(* LS Electric XG5000 project: Crane11 *)
(* PLC LSPLC *)
(* module base 0 slot 0: 입출력 모듈:XGH-DT4A (DC 24V 입력, 트랜지스터 출력 32점 ) *)
(* module base 0 slot 1: Cnet:XGL-C42A/B (Cnet 통신 모듈(RS-422/485, RS-422/485)) *)
VAR_GLOBAL
    AUTO_MODE_1 AT %IX0.0.0 : BOOL;
    AUTO_MODE_2 AT %IX0.0.1 : BOOL;
    AUTO_POSITION AT %IX0.0.6 : BOOL;
    AUTO_RESET AT %IX0.0.4 : BOOL;
    AUTO_RESUME AT %IX0.0.5 : BOOL;
    AUTO_START AT %IX0.0.2 : BOOL;
    AUTO_STOP AT %IX0.0.3 : BOOL;
    DRV_VAL AT %MW1 : WORD;
    DRV_VAL_GLOBAL : WORD;
    FREQ_VAL AT %MW0 : WORD;
    FREQ_VAL_GLOBAL : WORD;
    HALL_SENSOR_RPM AT %IX0.0.11 : BOOL;
    LED_AUTO_POSITION AT %QX0.0.19 : BOOL;
    LED_AUTO_RESET AT %QX0.0.20 : BOOL;
    LED_AUTO_RESUME AT %QX0.0.18 : BOOL;
    LED_AUTO_START AT %QX0.0.16 : BOOL;
    LED_AUTO_STOP AT %QX0.0.17 : BOOL;
    LIMITE_SW_BOTTOM_LEFT AT %IX0.0.13 : BOOL;
    LIMITE_SW_BOTTOM_RIGHT AT %IX0.0.15 : BOOL;
    LIMITE_SW_TOP_LEFT AT %IX0.0.12 : BOOL;
    LIMITE_SW_TOP_RIGHT AT %IX0.0.14 : BOOL;
    MODE_SELECT_AUTO AT %IX0.0.9 : BOOL;
    MODE_SELECT_PASSIVE AT %IX0.0.10 : BOOL;
    STATE_AUTO_MODE_1 : BOOL;
    STATE_AUTO_MODE_2 : BOOL;
    STATE_LIMITE_SW_BOTTOM_LEFT : BOOL;
    STATE_LIMITE_SW_BOTTOM_RIGHT : BOOL;
    STATE_POSITION : BOOL;
    STATE_RESET : BOOL;
    STATE_RESUME : BOOL;
    STATE_START : BOOL;
    STATE_STOP : BOOL;
    STATE_STOP_EMERGENCY : BOOL;
    STOP_EMERGENCY AT %IX0.0.7 : BOOL;
    SUCCESS_POSITION : BOOL;
    SUCCESS_RESET : BOOL;
    VAL_STATE_RESET : BOOL;
END_VAR

FUNCTION_BLOCK FB_LED_FLASH
(* 램프 점멸 동작 *)
VAR_INPUT
    EN_SW : BOOL;
    T_ON : TIME;
    T_OFF : TIME;
END_VAR
VAR_OUTPUT
    OUT_LAMP : BOOL;
END_VAR
VAR
    TIMER_1 : TON;
    TIMER_2 : TON;
END_VAR
(* 1. TIMER_1 동작: 시작 스위치가 켜져 있고, TIMER_2가 꺼져있을 때(.Q가 아닐 때) *)
TIMER_1(IN := EN_SW AND NOT TIMER_2.Q, PT := T_ON);

(* 2. TIMER_2 동작: TIMER_1이 완료되었을 때(.Q 일 때) *)
TIMER_2(IN := TIMER_1.Q, PT := T_OFF);

(* 3. 램프 출력: 스위치 ON 상태이고, TIMER_1이 도는 동안(아직 .Q가 안 떴을 때) *)
IF EN_SW AND NOT TIMER_1.Q THEN
    OUT_LAMP := TRUE;
ELSE
    OUT_LAMP := FALSE;
END_IF;
END_FUNCTION_BLOCK

FUNCTION_BLOCK FB_SELF_HOLD
VAR_INPUT
    START_SW : BOOL;
    STOP_SW : BOOL;
END_VAR
VAR_OUTPUT
    MOTOR_START : BOOL;
    MOTOR_STOP : BOOL;
END_VAR
IF STOP_SW THEN
    MOTOR_START := FALSE; // 실제 출력 변수 직접 제어
    MOTOR_STOP  := TRUE;
ELSIF START_SW THEN
    MOTOR_START := TRUE;
    MOTOR_STOP  := FALSE;
END_IF;
END_FUNCTION_BLOCK

PROGRAM LED_OUTPUT (* task: 스캔 프로그램 *)
(* LED출력관련 *)
VAR_EXTERNAL
    AUTO_POSITION : BOOL; (* AT %IX0.0.6 *)
    AUTO_RESET : BOOL; (* AT %IX0.0.4 *)
    AUTO_RESUME : BOOL; (* AT %IX0.0.5 *)
    AUTO_START : BOOL; (* AT %IX0.0.2 *)
    AUTO_STOP : BOOL; (* AT %IX0.0.3 *)
    LED_AUTO_POSITION : BOOL; (* AT %QX0.0.19 *)
    LED_AUTO_RESET : BOOL; (* AT %QX0.0.20 *)
    LED_AUTO_RESUME : BOOL; (* AT %QX0.0.18 *)
    LED_AUTO_START : BOOL; (* AT %QX0.0.16 *)
    LED_AUTO_STOP : BOOL; (* AT %QX0.0.17 *)
    STATE_POSITION : BOOL;
    STATE_RESET : BOOL;
    STATE_RESUME : BOOL;
    STATE_START : BOOL;
    STATE_STOP : BOOL;
    STATE_STOP_EMERGENCY : BOOL;
    STOP_EMERGENCY : BOOL; (* AT %IX0.0.7 *)
    SUCCESS_POSITION : BOOL;
    SUCCESS_RESET : BOOL;
END_VAR
VAR
    AUTO_RESET_STATE : BOOL;
    AUTO_STOP_STATE : BOOL;
    HOLD_EMERGENCY : FB_SELF_HOLD;
    HOLD_POSITION : FB_SELF_HOLD;
    HOLD_POSITION1 : FB_SELF_HOLD;
    HOLD_RESET : FB_SELF_HOLD;
    HOLD_RESET1 : FB_SELF_HOLD;
    HOLD_RESET2 : FB_SELF_HOLD;
    HOLD_START : FB_SELF_HOLD;
    HOLD_START1 : FB_SELF_HOLD;
    HOLD_START2 : FB_SELF_HOLD;
    HOLD_START3 : FB_SELF_HOLD;
    HOLD_STOP : FB_SELF_HOLD;
    LAMP_POSITION : FB_LED_FLASH;
    LAMP_RESET : FB_LED_FLASH;
    LAMP_RESUME : FB_LED_FLASH;
    LOCAL_POSITION : BOOL;
    LOCAL_RESET : BOOL;
    LOCAL_STOP_EMERGENCY : BOOL;
    RESET_STATE : BOOL;
    VAL_STATE : BOOL;
END_VAR

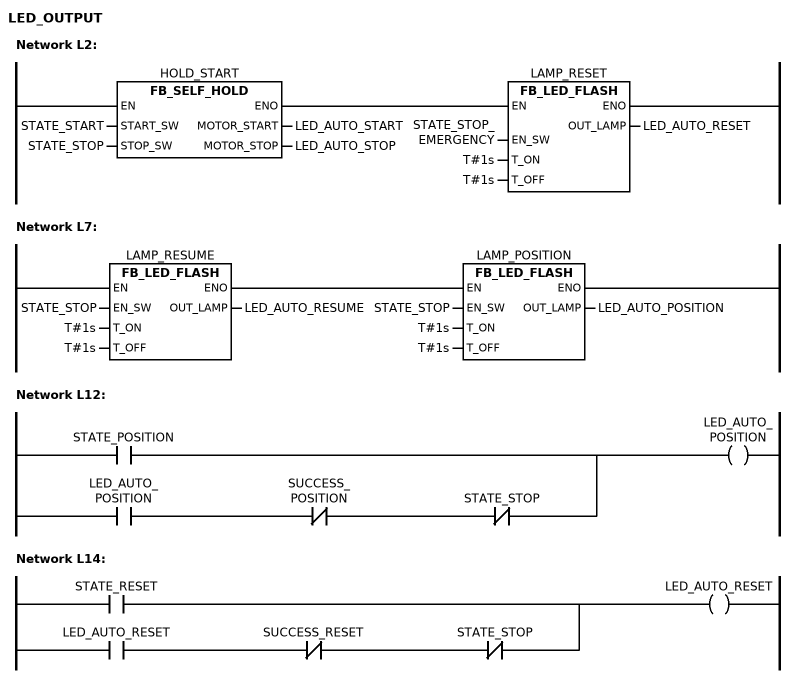
(* Rung L2 *)
HOLD_START(START_SW := STATE_START, STOP_SW := STATE_STOP, MOTOR_START => LED_AUTO_START, MOTOR_STOP => LED_AUTO_STOP);
LAMP_RESET(EN_SW := STATE_STOP_EMERGENCY, T_ON := T#1s, T_OFF := T#1s, OUT_LAMP => LED_AUTO_RESET);
(* Rung L7 *)
LAMP_RESUME(EN_SW := STATE_STOP, T_ON := T#1s, T_OFF := T#1s, OUT_LAMP => LED_AUTO_RESUME);
LAMP_POSITION(EN_SW := STATE_STOP, T_ON := T#1s, T_OFF := T#1s, OUT_LAMP => LED_AUTO_POSITION);
(* Rung L12 *)
LED_AUTO_POSITION := STATE_POSITION OR (LED_AUTO_POSITION AND NOT SUCCESS_POSITION AND NOT STATE_STOP);
(* Rung L14 *)
LED_AUTO_RESET := STATE_RESET OR (LED_AUTO_RESET AND NOT SUCCESS_RESET AND NOT STATE_STOP);
END_PROGRAM

PROGRAM AUTO_TIME (* task: 스캔 프로그램 *)
VAR_EXTERNAL
    AUTO_MODE_1 : BOOL; (* AT %IX0.0.0 *)
    AUTO_START : BOOL; (* AT %IX0.0.2 *)
    AUTO_STOP : BOOL; (* AT %IX0.0.3 *)
    MODE_SELECT_AUTO : BOOL; (* AT %IX0.0.9 *)
    STOP_EMERGENCY : BOOL; (* AT %IX0.0.7 *)
END_VAR
VAR
    COUNT_DOWN1 : TP;
    COUNT_DOWN2 : TP;
    DRV_VAL_LOCAL : WORD;
    FREQ_VAL_LOCAL : WORD;
    FREQ_VAL_START : WORD;
    IDLE : BOOL;
    INVERTER_STATE : BOOL;
    LOOP_SIGNAL : BOOL;
    RUN_FORWARD : BOOL;
    RUN_MOTOR : BOOL;
    RUN_REVERSE : BOOL;
    TARGET_TIME_FORWARD : TIME;
    TARGET_TIME_REVERSE : TIME;
    TIME_WAIT : TIME;
    VAL_DIV_FORWARD AT %MD151 : REAL := 1;
    VAL_DIV_REVERSE AT %MD152 : REAL := 1;
    VAL_Hz : REAL;
    VAL_MODE_FORWARD AT %MW11 : WORD := 2;
    VAL_MODE_REVERSE AT %MW12 : WORD := 4;
    VAL_MODE_WAIT : WORD;
    VAL_SPEED : WORD;
    VAL_TIME_DINT_FORWARD : DINT;
    VAL_TIME_DINT_REVERSE : DINT;
    VAL_TIME_REAL_FORWARD : REAL;
    VAL_TIME_REAL_REVERSE : REAL;
    VAL_TIME_UDINT_FORWARD : UDINT;
    VAL_TIME_UDINT_REVERSE : UDINT;
    대기1 : TON;
    대기2 : TON;
END_VAR
VAR
    _e1 : F_TRIG;
    _e2 : F_TRIG;
END_VAR

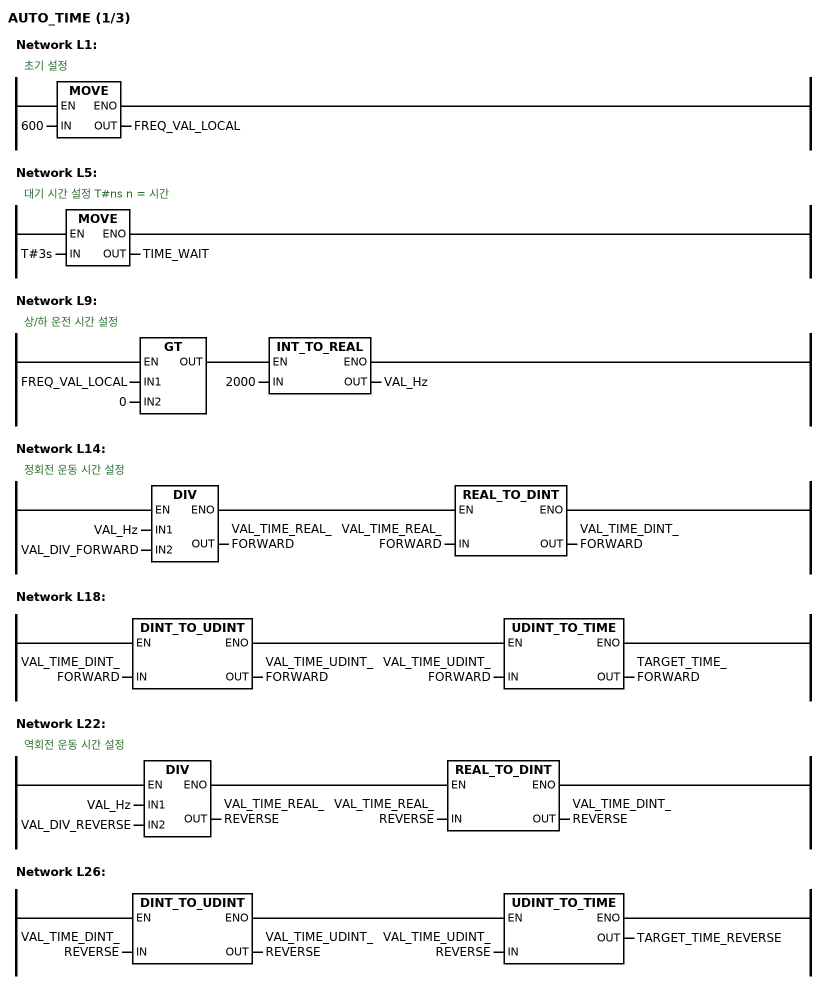
(* 초기 설정 *)
(* Rung L1 *)
FREQ_VAL_LOCAL := 600;
(* 대기 시간 설정 T#ns n = 시간 *)
(* Rung L5 *)
TIME_WAIT := T#3s;
(* 상/하 운전 시간 설정 *)
(* Rung L9 *)
IF FREQ_VAL_LOCAL > 0 THEN VAL_Hz := INT_TO_REAL(2000); END_IF;
(* 정회전 운동 시간 설정 *)
(* Rung L14 *)
VAL_TIME_REAL_FORWARD := VAL_Hz / VAL_DIV_FORWARD;
VAL_TIME_DINT_FORWARD := REAL_TO_DINT(VAL_TIME_REAL_FORWARD);
(* Rung L18 *)
VAL_TIME_UDINT_FORWARD := DINT_TO_UDINT(VAL_TIME_DINT_FORWARD);
TARGET_TIME_FORWARD := UDINT_TO_TIME(VAL_TIME_UDINT_FORWARD);
(* 역회전 운동 시간 설정 *)
(* Rung L22 *)
VAL_TIME_REAL_REVERSE := VAL_Hz / VAL_DIV_REVERSE;
VAL_TIME_DINT_REVERSE := REAL_TO_DINT(VAL_TIME_REAL_REVERSE);
(* Rung L26 *)
VAL_TIME_UDINT_REVERSE := DINT_TO_UDINT(VAL_TIME_DINT_REVERSE);
TARGET_TIME_REVERSE := UDINT_TO_TIME(VAL_TIME_UDINT_REVERSE);

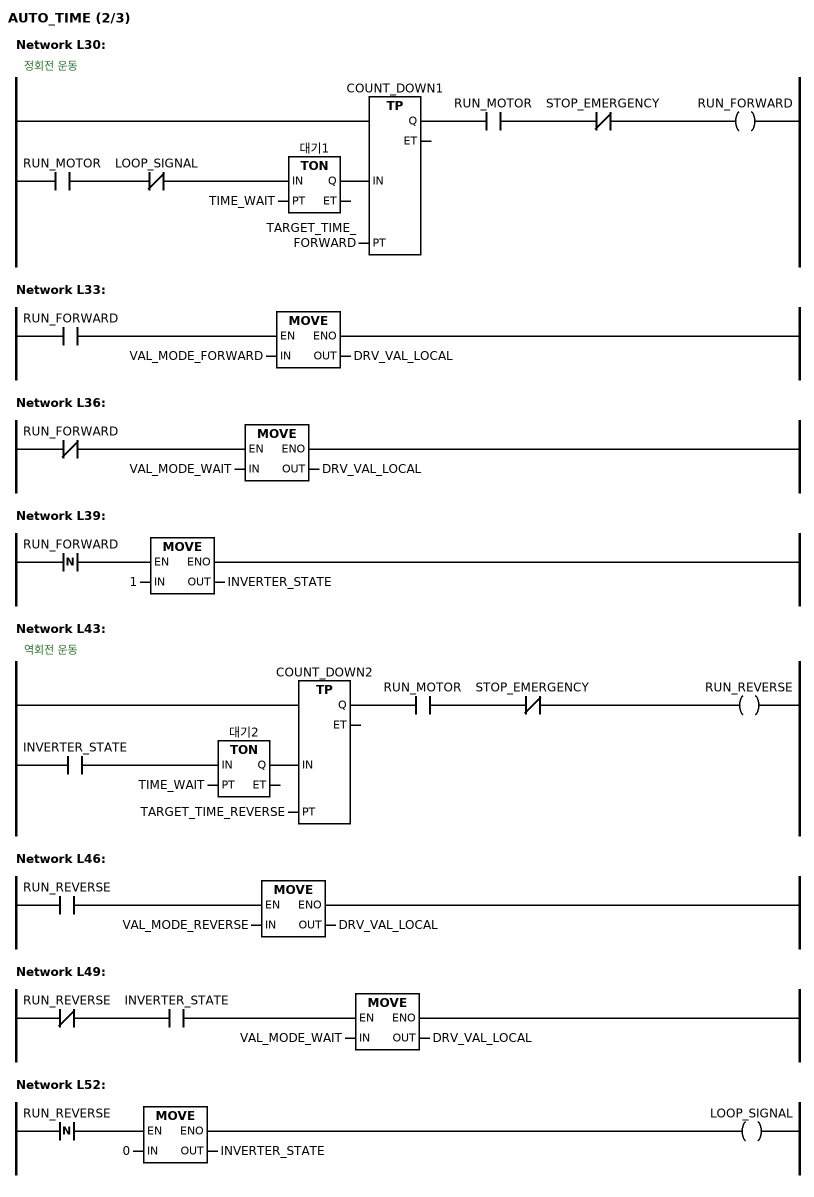
(* 정회전 운동 *)
(* Rung L30 *)
대기1(IN := RUN_MOTOR AND NOT LOOP_SIGNAL, PT := TIME_WAIT);
COUNT_DOWN1(IN := 대기1.Q, PT := TARGET_TIME_FORWARD);
RUN_FORWARD := COUNT_DOWN1.Q AND RUN_MOTOR AND NOT STOP_EMERGENCY;
(* Rung L33 *)
IF RUN_FORWARD THEN DRV_VAL_LOCAL := VAL_MODE_FORWARD; END_IF;
(* Rung L36 *)
IF NOT RUN_FORWARD THEN DRV_VAL_LOCAL := VAL_MODE_WAIT; END_IF;
(* Rung L39 *)
_e1(CLK := RUN_FORWARD);
IF _e1.Q THEN INVERTER_STATE := 1; END_IF;
(* 역회전 운동 *)
(* Rung L43 *)
대기2(IN := INVERTER_STATE, PT := TIME_WAIT);
COUNT_DOWN2(IN := 대기2.Q, PT := TARGET_TIME_REVERSE);
RUN_REVERSE := COUNT_DOWN2.Q AND RUN_MOTOR AND NOT STOP_EMERGENCY;
(* Rung L46 *)
IF RUN_REVERSE THEN DRV_VAL_LOCAL := VAL_MODE_REVERSE; END_IF;
(* Rung L49 *)
IF NOT RUN_REVERSE AND INVERTER_STATE THEN DRV_VAL_LOCAL := VAL_MODE_WAIT; END_IF;
(* Rung L52 *)
_e2(CLK := RUN_REVERSE);
IF _e2.Q THEN INVERTER_STATE := 0; END_IF;
LOOP_SIGNAL := _e2.Q;

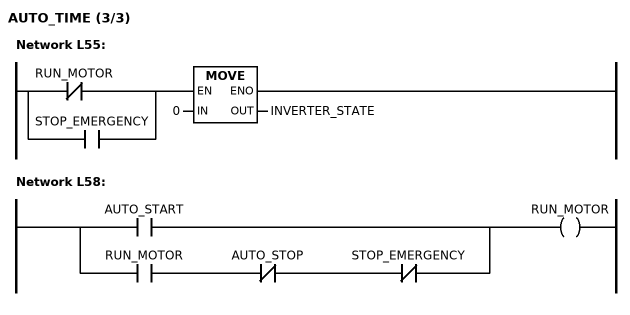
(* Rung L55 *)
IF NOT RUN_MOTOR OR STOP_EMERGENCY THEN INVERTER_STATE := 0; END_IF;
(* Rung L58 *)
RUN_MOTOR := AUTO_START OR (RUN_MOTOR AND NOT AUTO_STOP AND NOT STOP_EMERGENCY);
END_PROGRAM

PROGRAM INVERTER_CONTROL (* task: 스캔 프로그램 *)
VAR_EXTERNAL
    AUTO_MODE_1 : BOOL; (* AT %IX0.0.0 *)
    AUTO_MODE_2 : BOOL; (* AT %IX0.0.1 *)
    AUTO_STOP : BOOL; (* AT %IX0.0.3 *)
    DRV_VAL : WORD; (* AT %MW1 *)
    DRV_VAL_GLOBAL : WORD;
    FREQ_VAL : WORD; (* AT %MW0 *)
    FREQ_VAL_GLOBAL : WORD;
    STATE_POSITION : BOOL;
    STATE_RESET : BOOL;
    STATE_RESUME : BOOL;
    STATE_START : BOOL;
    STATE_STOP : BOOL;
    STATE_STOP_EMERGENCY : BOOL;
    STOP_EMERGENCY : BOOL; (* AT %IX0.0.7 *)
END_VAR
VAR
    DRV_VAL_LOCAL : WORD;
    FREQ_VAL_LOCAL : WORD;
    IDLE : BOOL;
    LIMITE_TRIGGER_BOTTOM : BOOL;
    LIMITE_TRIGGER_TOP : BOOL;
END_VAR

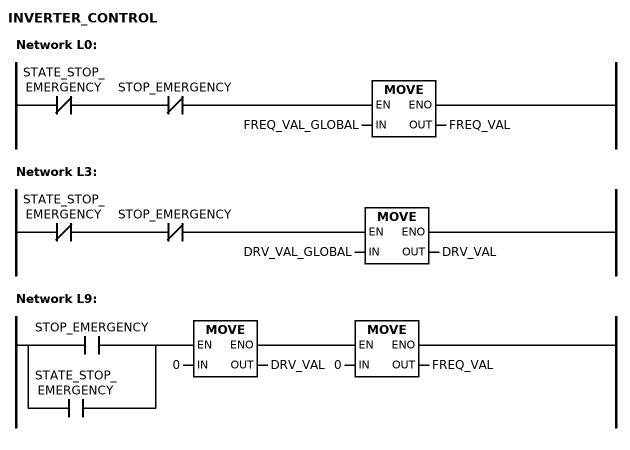
(* Rung L0 *)
IF NOT STATE_STOP_EMERGENCY AND NOT STOP_EMERGENCY THEN FREQ_VAL := FREQ_VAL_GLOBAL; END_IF;
(* Rung L3 *)
IF NOT STATE_STOP_EMERGENCY AND NOT STOP_EMERGENCY THEN DRV_VAL := DRV_VAL_GLOBAL; END_IF;
(* Rung L9 *)
IF STOP_EMERGENCY OR STATE_STOP_EMERGENCY THEN
    DRV_VAL := 0;
    FREQ_VAL := 0;
END_IF;
END_PROGRAM

PROGRAM RESET (* task: 스캔 프로그램 *)
VAR
    AUTO_RESET_STATE : BOOL;
    AUTO_RESUME_STATE : BOOL;
    COUNT_DOWN2 : TP;
    COUNT_DOWN3 : TP;
    COUNT_DOWN4 : TP;
    HOLD_FORWARD : FB_SELF_HOLD;
    VAL_STATE : BOOL;
    VAL_STATE_FORWARD : BOOL;
    VAL_STATE_IDLE : BOOL;
    VAL_STATE_REVERSE : BOOL;
    VAL_STATE_SUCCESS : BOOL;
END_VAR
VAR_EXTERNAL
    DRV_VAL_GLOBAL : WORD;
    FREQ_VAL_GLOBAL : WORD;
    LIMITE_SW_BOTTOM_LEFT : BOOL; (* AT %IX0.0.13 *)
    LIMITE_SW_BOTTOM_RIGHT : BOOL; (* AT %IX0.0.15 *)
    STATE_LIMITE_SW_BOTTOM_LEFT : BOOL;
    STATE_LIMITE_SW_BOTTOM_RIGHT : BOOL;
    STATE_POSITION : BOOL;
    STATE_RESET : BOOL;
    STATE_STOP : BOOL;
    SUCCESS_POSITION : BOOL;
    SUCCESS_RESET : BOOL;
    VAL_STATE_RESET : BOOL;
END_VAR
VAR
    _p1 : BOOL;
    _e2 : F_TRIG;
    _e3 : F_TRIG;
END_VAR

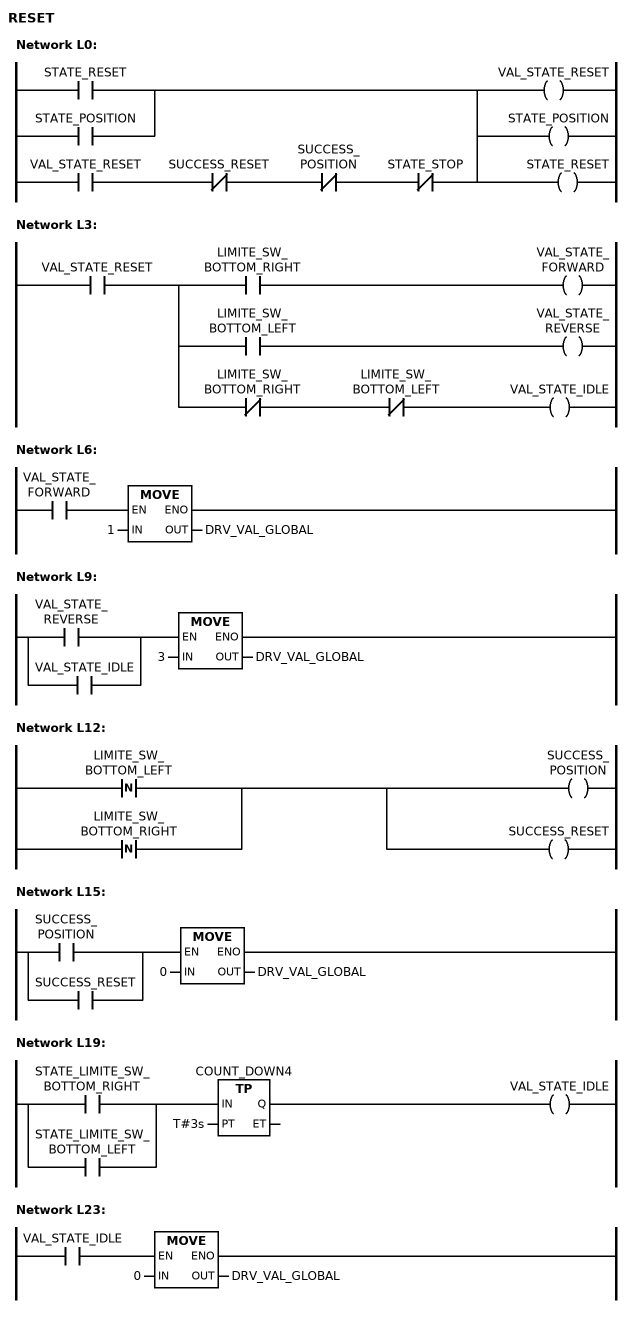
(* Rung L0 *)
_p1 := STATE_RESET OR STATE_POSITION OR (VAL_STATE_RESET AND NOT SUCCESS_RESET AND NOT SUCCESS_POSITION AND NOT STATE_STOP);
VAL_STATE_RESET := _p1;
STATE_POSITION := _p1;
STATE_RESET := _p1;
(* Rung L3 *)
VAL_STATE_FORWARD := VAL_STATE_RESET AND LIMITE_SW_BOTTOM_RIGHT;
VAL_STATE_REVERSE := VAL_STATE_RESET AND LIMITE_SW_BOTTOM_LEFT;
VAL_STATE_IDLE := VAL_STATE_RESET AND NOT LIMITE_SW_BOTTOM_RIGHT AND NOT LIMITE_SW_BOTTOM_LEFT;
(* Rung L6 *)
IF VAL_STATE_FORWARD THEN DRV_VAL_GLOBAL := 1; END_IF;
(* Rung L9 *)
IF VAL_STATE_REVERSE OR VAL_STATE_IDLE THEN DRV_VAL_GLOBAL := 3; END_IF;
(* Rung L12 *)
_e2(CLK := LIMITE_SW_BOTTOM_LEFT);
_e3(CLK := LIMITE_SW_BOTTOM_RIGHT);
SUCCESS_POSITION := _e2.Q OR _e3.Q;
SUCCESS_RESET := _e2.Q OR _e3.Q;
(* Rung L15 *)
IF SUCCESS_POSITION OR SUCCESS_RESET THEN DRV_VAL_GLOBAL := 0; END_IF;
(* Rung L19 *)
COUNT_DOWN4(IN := STATE_LIMITE_SW_BOTTOM_RIGHT OR STATE_LIMITE_SW_BOTTOM_LEFT, PT := T#3s);
VAL_STATE_IDLE := COUNT_DOWN4.Q;
(* Rung L23 *)
IF VAL_STATE_IDLE THEN DRV_VAL_GLOBAL := 0; END_IF;
END_PROGRAM

PROGRAM SW_CONTROL (* task: 스캔 프로그램 *)
VAR_EXTERNAL
    AUTO_MODE_1 : BOOL; (* AT %IX0.0.0 *)
    AUTO_MODE_2 : BOOL; (* AT %IX0.0.1 *)
    AUTO_POSITION : BOOL; (* AT %IX0.0.6 *)
    AUTO_RESET : BOOL; (* AT %IX0.0.4 *)
    AUTO_RESUME : BOOL; (* AT %IX0.0.5 *)
    AUTO_START : BOOL; (* AT %IX0.0.2 *)
    AUTO_STOP : BOOL; (* AT %IX0.0.3 *)
    LED_AUTO_POSITION : BOOL; (* AT %QX0.0.19 *)
    LED_AUTO_RESET : BOOL; (* AT %QX0.0.20 *)
    LIMITE_SW_BOTTOM_LEFT : BOOL; (* AT %IX0.0.13 *)
    LIMITE_SW_BOTTOM_RIGHT : BOOL; (* AT %IX0.0.15 *)
    LIMITE_SW_TOP_LEFT : BOOL; (* AT %IX0.0.12 *)
    LIMITE_SW_TOP_RIGHT : BOOL; (* AT %IX0.0.14 *)
    STATE_AUTO_MODE_1 : BOOL;
    STATE_AUTO_MODE_2 : BOOL;
    STATE_LIMITE_SW_BOTTOM_LEFT : BOOL;
    STATE_LIMITE_SW_BOTTOM_RIGHT : BOOL;
    STATE_POSITION : BOOL;
    STATE_RESET : BOOL;
    STATE_RESUME : BOOL;
    STATE_START : BOOL;
    STATE_STOP : BOOL;
    STATE_STOP_EMERGENCY : BOOL;
    STOP_EMERGENCY : BOOL; (* AT %IX0.0.7 *)
    SUCCESS_POSITION : BOOL;
    SUCCESS_RESET : BOOL;
END_VAR
VAR
    HOLD_EMERGENCY : FB_SELF_HOLD;
    HOLD_POSITION : FB_SELF_HOLD;
    HOLD_RESET : FB_SELF_HOLD;
    HOLD_RESET1 : FB_SELF_HOLD;
END_VAR

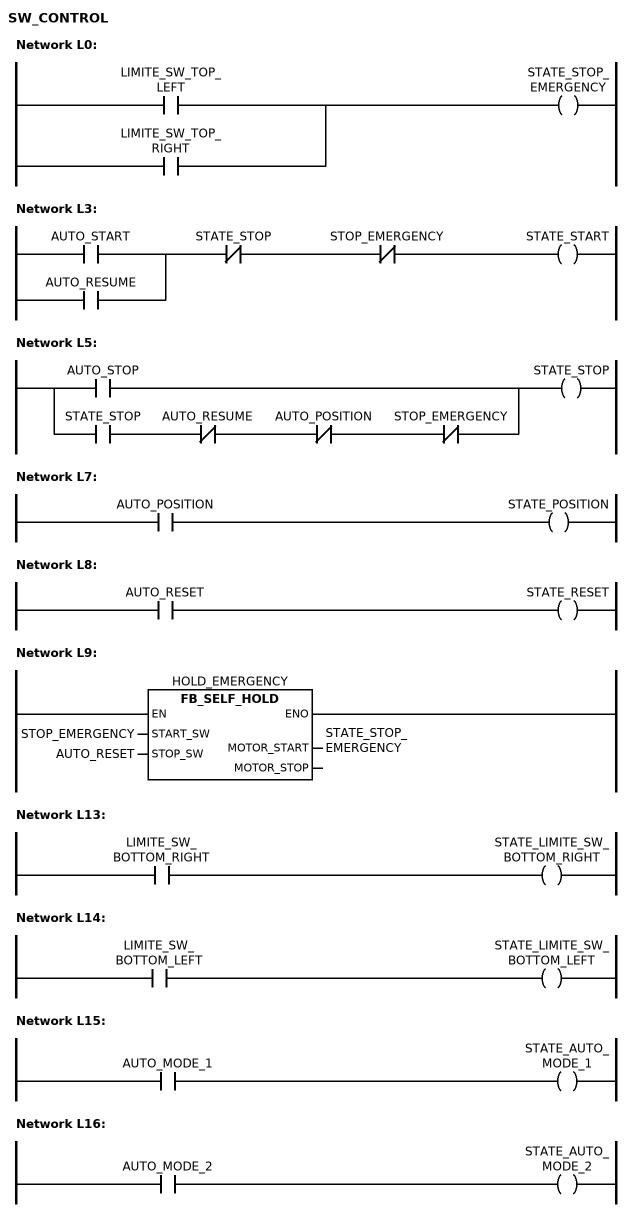
(* Rung L0 *)
STATE_STOP_EMERGENCY := LIMITE_SW_TOP_LEFT OR LIMITE_SW_TOP_RIGHT;
(* Rung L3 *)
STATE_START := (AUTO_START OR AUTO_RESUME) AND NOT STATE_STOP AND NOT STOP_EMERGENCY;
(* Rung L5 *)
STATE_STOP := AUTO_STOP OR (STATE_STOP AND NOT AUTO_RESUME AND NOT AUTO_POSITION AND NOT STOP_EMERGENCY);
(* Rung L7 *)
STATE_POSITION := AUTO_POSITION;
(* Rung L8 *)
STATE_RESET := AUTO_RESET;
(* Rung L9 *)
HOLD_EMERGENCY(START_SW := STOP_EMERGENCY, STOP_SW := AUTO_RESET, MOTOR_START => STATE_STOP_EMERGENCY);
(* Rung L13 *)
STATE_LIMITE_SW_BOTTOM_RIGHT := LIMITE_SW_BOTTOM_RIGHT;
(* Rung L14 *)
STATE_LIMITE_SW_BOTTOM_LEFT := LIMITE_SW_BOTTOM_LEFT;
(* Rung L15 *)
STATE_AUTO_MODE_1 := AUTO_MODE_1;
(* Rung L16 *)
STATE_AUTO_MODE_2 := AUTO_MODE_2;
END_PROGRAM

PROGRAM AUTO_SW (* task: 스캔 프로그램 *)
VAR
    COUNT_DOWN2 : TP;
    HOLD_START : FB_SELF_HOLD;
    TARGET_TIME_REVERSE : TIME;
    TIME_WAIT : TIME;
    VAL_STATE : BOOL;
    VAL_STATE_FORWARD : BOOL;
    VAL_STATE_IDLE : BOOL;
    VAL_STATE_IDLE_LOCAL : BOOL;
    VAL_STATE_REVERSE : BOOL;
    WAIT : TON;
    대기1 : TON;
END_VAR
VAR_EXTERNAL
    DRV_VAL_GLOBAL : WORD;
    LIMITE_SW_BOTTOM_LEFT : BOOL; (* AT %IX0.0.13 *)
    LIMITE_SW_BOTTOM_RIGHT : BOOL; (* AT %IX0.0.15 *)
    STATE_LIMITE_SW_BOTTOM_LEFT : BOOL;
    STATE_LIMITE_SW_BOTTOM_RIGHT : BOOL;
    STATE_POSITION : BOOL;
    STATE_RESET : BOOL;
    STATE_START : BOOL;
    STATE_STOP : BOOL;
    SUCCESS_POSITION : BOOL;
    SUCCESS_RESET : BOOL;
    VAL_STATE_RESET : BOOL;
END_VAR

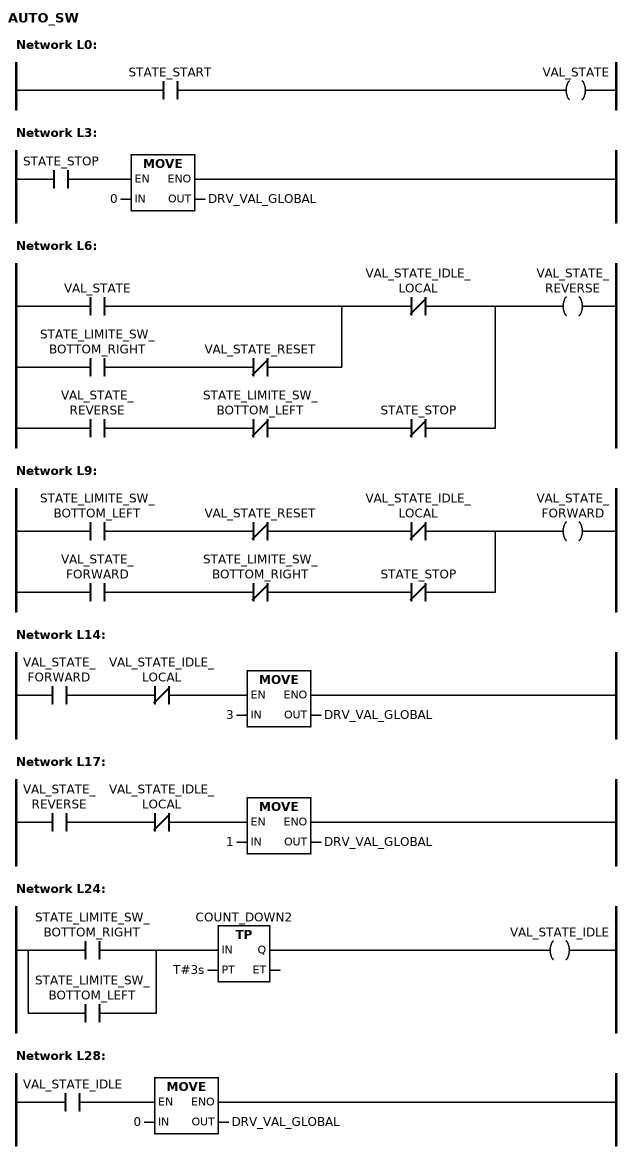
(* Rung L0 *)
VAL_STATE := STATE_START;
(* Rung L3 *)
IF STATE_STOP THEN DRV_VAL_GLOBAL := 0; END_IF;
(* Rung L6 *)
VAL_STATE_REVERSE := ((VAL_STATE OR (STATE_LIMITE_SW_BOTTOM_RIGHT AND NOT VAL_STATE_RESET)) AND NOT VAL_STATE_IDLE_LOCAL) OR (VAL_STATE_REVERSE AND NOT STATE_LIMITE_SW_BOTTOM_LEFT AND NOT STATE_STOP);
(* Rung L9 *)
VAL_STATE_FORWARD := (STATE_LIMITE_SW_BOTTOM_LEFT AND NOT VAL_STATE_RESET AND NOT VAL_STATE_IDLE_LOCAL) OR (VAL_STATE_FORWARD AND NOT STATE_LIMITE_SW_BOTTOM_RIGHT AND NOT STATE_STOP);
(* Rung L14 *)
IF VAL_STATE_FORWARD AND NOT VAL_STATE_IDLE_LOCAL THEN DRV_VAL_GLOBAL := 3; END_IF;
(* Rung L17 *)
IF VAL_STATE_REVERSE AND NOT VAL_STATE_IDLE_LOCAL THEN DRV_VAL_GLOBAL := 1; END_IF;
(* Rung L24 *)
COUNT_DOWN2(IN := STATE_LIMITE_SW_BOTTOM_RIGHT OR STATE_LIMITE_SW_BOTTOM_LEFT, PT := T#3s);
VAL_STATE_IDLE := COUNT_DOWN2.Q;
(* Rung L28 *)
IF VAL_STATE_IDLE THEN DRV_VAL_GLOBAL := 0; END_IF;
END_PROGRAM

PROGRAM AUTO_Hz (* task: 스캔 프로그램 *)
VAR_EXTERNAL
    FREQ_VAL_GLOBAL : WORD;
    STATE_AUTO_MODE_1 : BOOL;
    STATE_AUTO_MODE_2 : BOOL;
END_VAR
VAR
    FREQ_VAL_LOCAL : WORD;
END_VAR

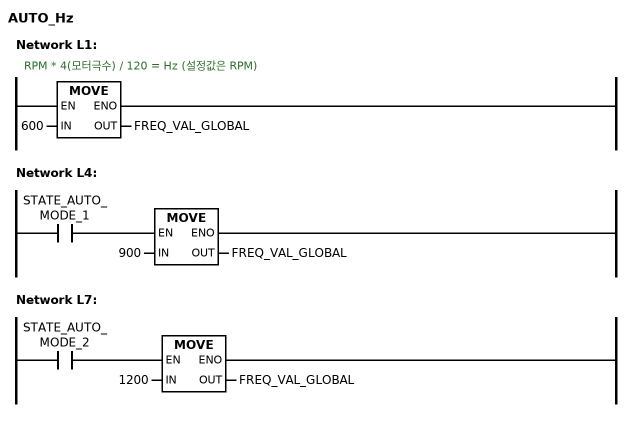
(* RPM * 4(모터극수) / 120 = Hz (설정값은 RPM) *)
(* Rung L1 *)
FREQ_VAL_GLOBAL := 600;
(* Rung L4 *)
IF STATE_AUTO_MODE_1 THEN FREQ_VAL_GLOBAL := 900; END_IF;
(* Rung L7 *)
IF STATE_AUTO_MODE_2 THEN FREQ_VAL_GLOBAL := 1200; END_IF;
END_PROGRAM